FUNCTION_BLOCK logiBUS_AI_MV (* Input service interface function block for analog input in millivolts *)
  (* Description: Copyright (c) 2017 fortiss GmbH, HR Agrartechnik GmbH This program and the accompanying materials are made available under the terms of the Eclipse Public License 2.0 which is available at https://www.eclipse.org/legal/epl-2.0/ SPDX-License-Identifier: EPL-2.0 AnalogInput_hysteresis = 0 switches the change trigger off (use 1 to see every change). TimeDelta = 0 or 16#FFFFFFFF switches the cyclic IND off. With both off the block sends no IND (value only via REQ). IN = calibrated voltage at the pin in mV (ADC calibration of the chip from eFuse, attenuation as for logiBUS_AI_ID: ESP32-S3 about 0-2900 mV, ESP32-P4 about 0-3300 mV). Without calibration for the channel (e.g. ESP32-S31 with the current ESP-IDF) INIT fails with STATUS = 'ADC calibration not available'. *)
  (* Version 1.0, 2026-11-13, Franz Höpfinger, HR Agrartechnik GmbH *)
  PACKAGE logiBUS::io::AI;
  (* Documentation:
  logiBUS_AI_MV
   🇩🇪 Deutsch
   Service-Interface-Funktionsblock für einen analogen Eingang in Millivolt. Wie logiBUS_AI_ID, aber IN liefert die kalibrierte Spannung am Pin statt des Rohwerts.
   Wert von IN
   IN ist die Spannung am Pin des Chips in Millivolt (DWORD). Die Firmware rechnet den gemittelten Rohwert mit der Kalibrierung des Chips um (ESP-IDF adc_cali, Werte aus dem eFuse). Die Dämpfung ist dieselbe wie bei logiBUS_AI_ID: ESP32-S3 etwa 0-2900 mV (±50 mV), ESP32-P4 etwa 0-3300 mV (±15 mV), laut Datenblatt.
   Die Spannung an der Klemme hängt vom Spannungsteiler der Platine ab und ist nicht eingerechnet.
   Gibt es für den Kanal keine Kalibrierung (z. B. ESP32-S31 mit dem aktuellen ESP-IDF), meldet INIT QO = FALSE und STATUS = ADC calibration not available.
   Hysterese und Zeitsteuerung
   Wie bei logiBUS_AI_ID, aber AnalogInput_hysteresis gilt in mV.
   🇬🇧 English
   Service interface function block for one analog input in millivolts. Like logiBUS_AI_ID, but IN delivers the calibrated voltage at the pin instead of the raw value.
   Value of IN
   IN is the voltage at the chip pin in millivolts (DWORD). The firmware converts the averaged raw value with the chip calibration (ESP-IDF adc_cali, eFuse values). The attenuation is the same as for logiBUS_AI_ID: ESP32-S3 about 0-2900 mV (±50 mV), ESP32-P4 about 0-3300 mV (±15 mV), according to the datasheet.
   The voltage at the terminal depends on the voltage divider of the board and is not included.
   Without a calibration for the channel (e.g. ESP32-S31 with the current ESP-IDF), INIT returns QO = FALSE and STATUS = ADC calibration not available.
   Hysteresis and timing
   As for logiBUS_AI_ID, but AnalogInput_hysteresis is in mV.
  *)
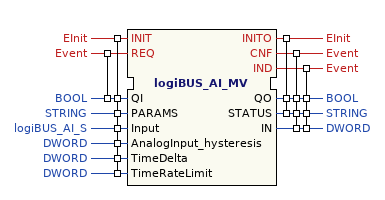
  EVENT_INPUT
    INIT : EInit WITH QI, PARAMS, Input, AnalogInput_hysteresis, TimeDelta, TimeRateLimit; (* Service Initialization *)
    REQ WITH QI; (* Service Request *)
  END_EVENT
  EVENT_OUTPUT
    INITO : EInit WITH QO, STATUS; (* Initialization Confirm *)
    CNF WITH QO, STATUS, IN; (* Confirmation of Requested Service *)
    IND WITH QO, STATUS, IN; (* Indication from Resource *)
  END_EVENT
  VAR_INPUT
    QI : BOOL; (* Event Input Qualifier *)
    PARAMS : STRING; (* Service Parameters *)
    Input : logiBUS::io::AI::logiBUS_AI_S := logiBUS_AI::Invalid; (* Identify the Input Input_I1..I8 *)
    AnalogInput_hysteresis : DWORD; (* IND when the voltage changes by more than this many mV (0 = off) *)
    TimeDelta : DWORD := 250; (* After How many ms an IND (poll interval, 0 or 16#FFFFFFFF = off) *)
    TimeRateLimit : DWORD := 100; (* Maximum 1 IND in how many ms. (< delta) *)
  END_VAR
  VAR_OUTPUT
    QO : BOOL; (* Event Output Qualifier *)
    STATUS : STRING; (* Service Status *)
    IN : DWORD; (* Input data from resource, calibrated voltage at the pin in mV *)
  END_VAR
END_FUNCTION_BLOCK
